Fanuc KAREL source: kt00135.KL

-- PROVISIONAL review KL for V1013-1; original PC SHA256 4c6c51d706d3555d31adc98a216263b64bacee091bf7303f48b7b7fd34232ec9
-- Incomplete behavior may be omitted. Consult companion uncertainty JSON. Do not deploy.
PROGRAM KT00135
%NOLOCKGROUP
VAR
  I1 : INTEGER
  OUT : INTEGER
-- UNRESOLVED_DECL H2 type=002017
BEGIN
  -- UNRESOLVED_PC offsets 5-16; opcodes 2E,23
  -- UNRESOLVED_PC offsets 21-35; opcodes 2E,22,9D,33,B4
  -- UNRESOLVED_PC offsets 40-62; opcodes 21,22,9D,33,B3,55,23
  -- UNRESOLVED_PC offsets 67-71; opcodes 7F
END KT00135
